Fanuc KAREL source: kd00017.KL

-- PROVISIONAL review KL for V940-1; original PC SHA256 ffe0f540755ae5a331bd5d33f45c77edb949f3d3b2d673eaac4cfbdf272d6a47
-- Incomplete behavior may be omitted. Consult companion uncertainty JSON. Do not deploy.
PROGRAM KD00017
%NOLOCKGROUP
VAR
  I : INTEGER
  J : INTEGER
  B : BOOLEAN
  R : REAL
  S : STRING[80]
BEGIN
  -- V9_ZERO_TABLE_METADATA_HINT layout=0001; no indexed target words; source/name/runtime held
  -- UNRESOLVED_PC offsets 5-12; opcodes 9C,23
  -- UNRESOLVED_PC offsets 17-24; opcodes 22,62
  -- UNRESOLVED_PC offsets 29-36; opcodes 22,28
  -- UNRESOLVED_PC offsets 41-45; opcodes 7F
END KD00017
